Yaskawa INFORM job: DROP.JBI

/JOB
//NAME DROP
//POS
///NPOS 0,0,0,4,0,0
///TOOL 0
///POSTYPE BASE
///RECTAN
///RCONF 0,0,0,0,0,0,0,0
P0008=0.000,0.000,300.000,0.00,0.00,0.00
P0009=0.000,-1332.000,600.000,180.00,0.00,0.00
P0010=0.000,-1332.000,390.000,180.00,0.00,0.00
P0011=0.000,0.000,200.000,0.00,0.00,0.00
//INST
///DATE 2026/10/27 16:49
///ATTR SC,RW
///GROUP1 RB1
NOP
SET B090 0
IMOV P008 V=I000 PL=0 BF DEC=50
MOVL P009 V=I000 PL=0 DEC=50
SET B090 1
MOVL P010 V=I000 PL=0 DEC=50
HAND HNO: 2 OFF
TIMER T=1.00
IMOV P011 V=I000 PL=0
END
